(* IEC 61131-3 sources: plc-workbench/customers/naidis-metall/magazine-swivel/plc/src, 2 files *)

(* ---- plant_sim.st ---- *)
(* Plant model of the magazine and swivel station, for the sim target only.
   Reads the valve coils and writes the sensors, once per 10 ms scan before Station.
   Positions count scans: one count per scan, so 40 counts = 400 ms of travel. *)

PROGRAM PlantSim
    VAR_EXTERNAL
        MAG_CylExtended : BOOL;
        MAG_CylRetracted : BOOL;
        GRP_PartGripped : BOOL;
        SWV_AtPickup : BOOL;
        SWV_AtDropdown : BOOL;
        MAG_PickupOccupied : BOOL;
        MAG_CylRetract : BOOL;
        GRP_Grip : BOOL;
        GRP_Release : BOOL;
        SWV_ToPickup : BOOL;
        SWV_ToDropdown : BOOL;
        SIM_PartsInMagazine : INT;
        SIM_PartsDelivered : INT;
        SIM_PartsLost : INT;
        SIM_VacuumFault : BOOL;
        SIM_SwivelJam : BOOL;
        SIM_SorterBlocked : BOOL;
        LNK_NextReady : BOOL;
    END_VAR
    VAR CONSTANT
        MagStroke : INT := 40;    (* 0 = extended, MagStroke = retracted *)
        SwvStroke : INT := 50;    (* 0 = at dropdown, SwvStroke = at pickup *)
        SortScans : INT := 100;   (* the sorter takes a delivered part away in 1 s *)
    END_VAR
    VAR
        MagPos : INT := 0;
        SwvPos : INT := 0;
        PartInFront : BOOL;       (* dropped from the magazine in front of the retracted cylinder *)
        PartAtPickup : BOOL;
        PartOnGripper : BOOL;
        Vacuum : BOOL;
        VacuumBuildUp : TON;
        SortCount : INT := 0;     (* > 0 while the sorter is busy with the last part *)
    END_VAR

    (* 1A1 magazine cylinder: 5/2 single solenoid, coil on retracts, spring extends *)
    IF MAG_CylRetract THEN
        IF MagPos < MagStroke THEN MagPos := MagPos + 1; END_IF;
    ELSIF MagPos > 0 THEN
        MagPos := MagPos - 1;
    END_IF;
    IF MagPos = MagStroke AND NOT PartInFront AND SIM_PartsInMagazine > 0 THEN
        PartInFront := TRUE;
        SIM_PartsInMagazine := SIM_PartsInMagazine - 1;
    END_IF;
    IF MagPos = 0 AND PartInFront THEN
        PartInFront := FALSE;
        PartAtPickup := TRUE;
    END_IF;

    (* 3A1 swivel: 5/3 closed centre, stops with both coils off or both on *)
    IF NOT SIM_SwivelJam THEN
        IF SWV_ToPickup AND NOT SWV_ToDropdown AND SwvPos < SwvStroke THEN
            SwvPos := SwvPos + 1;
        ELSIF SWV_ToDropdown AND NOT SWV_ToPickup AND SwvPos > 0 THEN
            SwvPos := SwvPos - 1;
        END_IF;
    END_IF;

    (* 2A1 vacuum gripper: valve keeps its last coil *)
    IF GRP_Grip AND NOT GRP_Release THEN
        Vacuum := TRUE;
    ELSIF GRP_Release AND NOT GRP_Grip THEN
        Vacuum := FALSE;
    END_IF;
    IF Vacuum AND SwvPos = SwvStroke AND PartAtPickup THEN
        PartAtPickup := FALSE;
        PartOnGripper := TRUE;
    END_IF;
    IF PartOnGripper AND (NOT Vacuum OR SIM_VacuumFault) THEN
        PartOnGripper := FALSE;
        IF SwvPos = 0 AND LNK_NextReady THEN
            SIM_PartsDelivered := SIM_PartsDelivered + 1;
            SortCount := SortScans;
        ELSIF SwvPos = 0 THEN
            SIM_PartsLost := SIM_PartsLost + 1;      (* dropped onto a sorter that was not ready *)
        ELSIF SwvPos = SwvStroke THEN
            PartAtPickup := TRUE;
        ELSE
            SIM_PartsLost := SIM_PartsLost + 1;
        END_IF;
    END_IF;
    VacuumBuildUp(IN := Vacuum AND PartOnGripper, PT := T#100MS);

    (* colour sorter downstream: ready over the IR link unless busy or blocked *)
    IF SortCount > 0 THEN SortCount := SortCount - 1; END_IF;

    MAG_CylExtended := MagPos = 0;
    MAG_CylRetracted := MagPos = MagStroke;
    MAG_PickupOccupied := PartAtPickup;
    SWV_AtDropdown := SwvPos = 0;
    SWV_AtPickup := SwvPos = SwvStroke;
    GRP_PartGripped := VacuumBuildUp.Q;
    LNK_NextReady := SortCount = 0 AND NOT SIM_SorterBlocked;
END_PROGRAM

(* ---- station.st ---- *)
(* Magazine and swivel station: step sequence.
   Spec: ../magazine-swivel.spec.md, section 5.
   I/O symbols are globals declared by the target (targets/*.st). *)

TYPE
    StepT : (
        S0_Ready,
        S1_MagRetract,
        S2_MagPushOut,
        S3_SwvToPickup,
        S4_VacuumOn,
        S5_WaitNextReady,
        S6_SwvToDropdown,
        S7_VacuumOff,
        S8_CycleEnd,
        S9_MagEmpty,
        S90_HomingRequired,
        S91_HomeSwivel,
        S92_HomeVacuumOff,
        S99_Alarm);
END_TYPE

PROGRAM Station
    VAR_EXTERNAL
        PNL_StartButton : BOOL;
        PNL_StopReleased : BOOL;
        PNL_Manual : BOOL;
        PNL_ResetButton : BOOL;
        PNL_EStopOk : BOOL;
        MAG_CylExtended : BOOL;
        MAG_CylRetracted : BOOL;
        GRP_PartGripped : BOOL;
        SWV_AtPickup : BOOL;
        SWV_AtDropdown : BOOL;
        MAG_PickupOccupied : BOOL;
        LNK_NextReady : BOOL;
        PNL_StartLamp : BOOL;
        PNL_ResetLamp : BOOL;
        PNL_LampQ1 : BOOL;
        PNL_LampQ2 : BOOL;
        MAG_CylRetract : BOOL;
        GRP_Grip : BOOL;
        GRP_Release : BOOL;
        SWV_ToPickup : BOOL;
        SWV_ToDropdown : BOOL;
        StepNo : INT;   (* Step as a number (S90 = 90) for HMI and simulation *)
    END_VAR
    VAR
        CurStep : StepT := S90_HomingRequired;
        LastStep : StepT := S90_HomingRequired;
        StepTimer : TON;
        StepTime : TIME;
        FirstScan : BOOL := TRUE;
        StartTrig : R_TRIG;
        ResetTrig : R_TRIG;
        StartP : BOOL;
        ResetP : BOOL;
        BlinkTimer : TON;
        Blink1Hz : BOOL;
        Home : BOOL;
        StopReq : BOOL;
    END_VAR

    StepTimer(IN := CurStep = LastStep, PT := T#24H);  (* restarts on every step change *)
    StepTime := StepTimer.ET;
    LastStep := CurStep;

    BlinkTimer(IN := NOT BlinkTimer.Q, PT := T#500MS);
    IF BlinkTimer.Q THEN Blink1Hz := NOT Blink1Hz; END_IF;

    StartTrig(CLK := PNL_StartButton);
    StartP := StartTrig.Q;
    ResetTrig(CLK := PNL_ResetButton);
    ResetP := ResetTrig.Q;

    Home := MAG_CylExtended AND SWV_AtDropdown;

    IF CurStep = S0_Ready OR CurStep = S9_MagEmpty THEN
        StopReq := FALSE;
    ELSIF NOT PNL_StopReleased THEN
        StopReq := TRUE;
    END_IF;

    IF FirstScan THEN
        IF Home THEN CurStep := S0_Ready; ELSE CurStep := S90_HomingRequired; END_IF;
    ELSIF NOT PNL_EStopOk THEN
        CurStep := S90_HomingRequired;
    ELSE
        CASE CurStep OF
        S90_HomingRequired:
            IF ResetP AND PNL_EStopOk THEN CurStep := S91_HomeSwivel; END_IF;

        S91_HomeSwivel:
            IF SWV_AtDropdown THEN CurStep := S92_HomeVacuumOff;
            ELSIF StepTime >= T#3S THEN CurStep := S99_Alarm; END_IF;

        S92_HomeVacuumOff:
            IF StepTime >= T#50MS AND Home THEN CurStep := S0_Ready;
            ELSIF StepTime >= T#3S THEN CurStep := S99_Alarm; END_IF;

        S0_Ready:
            IF NOT Home THEN CurStep := S90_HomingRequired;
            ELSIF StartP AND PNL_StopReleased THEN
                IF MAG_PickupOccupied THEN CurStep := S3_SwvToPickup; ELSE CurStep := S1_MagRetract; END_IF;
            END_IF;

        S1_MagRetract:
            IF MAG_CylRetracted THEN CurStep := S2_MagPushOut;
            ELSIF StepTime >= T#3S THEN CurStep := S99_Alarm; END_IF;

        S2_MagPushOut:
            IF MAG_CylExtended THEN
                IF MAG_PickupOccupied THEN CurStep := S3_SwvToPickup; ELSE CurStep := S9_MagEmpty; END_IF;
            ELSIF StepTime >= T#3S THEN CurStep := S99_Alarm; END_IF;

        S3_SwvToPickup:
            IF SWV_AtPickup THEN CurStep := S4_VacuumOn;
            ELSIF StepTime >= T#3S THEN CurStep := S99_Alarm; END_IF;

        S4_VacuumOn:
            IF GRP_PartGripped THEN CurStep := S5_WaitNextReady;
            ELSIF StepTime >= T#3S THEN CurStep := S99_Alarm; END_IF;  (* part not gripped *)

        S5_WaitNextReady:
            IF NOT GRP_PartGripped THEN CurStep := S99_Alarm;          (* part lost *)
            ELSIF LNK_NextReady THEN CurStep := S6_SwvToDropdown; END_IF;

        S6_SwvToDropdown:
            IF NOT GRP_PartGripped THEN CurStep := S99_Alarm;          (* part lost *)
            ELSIF SWV_AtDropdown THEN CurStep := S7_VacuumOff;
            ELSIF StepTime >= T#3S THEN CurStep := S99_Alarm; END_IF;

        S7_VacuumOff:
            IF StepTime >= T#50MS THEN CurStep := S8_CycleEnd; END_IF;

        S8_CycleEnd:
            IF StopReq OR PNL_Manual THEN CurStep := S0_Ready; ELSE CurStep := S1_MagRetract; END_IF;

        S9_MagEmpty:
            IF NOT Home THEN CurStep := S90_HomingRequired;
            ELSIF StartP AND PNL_StopReleased THEN CurStep := S1_MagRetract; END_IF;

        S99_Alarm:
            IF ResetP AND PNL_EStopOk THEN CurStep := S91_HomeSwivel; END_IF;
        END_CASE;
    END_IF;

    (* one line per output; never assigned anywhere else *)
    MAG_CylRetract := CurStep = S1_MagRetract AND SWV_AtDropdown;
    GRP_Grip := CurStep = S4_VacuumOn OR CurStep = S5_WaitNextReady OR CurStep = S6_SwvToDropdown;
    GRP_Release := CurStep = S92_HomeVacuumOff OR CurStep = S7_VacuumOff;
    SWV_ToPickup := (CurStep = S3_SwvToPickup OR CurStep = S4_VacuumOn OR CurStep = S5_WaitNextReady)
        AND MAG_CylExtended;
    SWV_ToDropdown := CurStep = S91_HomeSwivel OR CurStep = S92_HomeVacuumOff
        OR CurStep = S6_SwvToDropdown OR CurStep = S7_VacuumOff;
    PNL_StartLamp := (CurStep = S0_Ready OR CurStep = S9_MagEmpty) AND Blink1Hz
        OR CurStep = S1_MagRetract OR CurStep = S2_MagPushOut OR CurStep = S3_SwvToPickup
        OR CurStep = S4_VacuumOn OR CurStep = S5_WaitNextReady OR CurStep = S6_SwvToDropdown
        OR CurStep = S7_VacuumOff OR CurStep = S8_CycleEnd;
    PNL_ResetLamp := CurStep = S90_HomingRequired AND (Blink1Hz OR NOT PNL_EStopOk)
        OR CurStep = S91_HomeSwivel OR CurStep = S92_HomeVacuumOff
        OR CurStep = S99_Alarm AND Blink1Hz;
    PNL_LampQ1 := PNL_ResetLamp;   (* same steps and modifiers as the reset lamp *)
    PNL_LampQ2 := PNL_ResetLamp OR CurStep = S9_MagEmpty AND Blink1Hz;

    CASE CurStep OF
    S0_Ready: StepNo := 0;
    S1_MagRetract: StepNo := 1;
    S2_MagPushOut: StepNo := 2;
    S3_SwvToPickup: StepNo := 3;
    S4_VacuumOn: StepNo := 4;
    S5_WaitNextReady: StepNo := 5;
    S6_SwvToDropdown: StepNo := 6;
    S7_VacuumOff: StepNo := 7;
    S8_CycleEnd: StepNo := 8;
    S9_MagEmpty: StepNo := 9;
    S90_HomingRequired: StepNo := 90;
    S91_HomeSwivel: StepNo := 91;
    S92_HomeVacuumOff: StepNo := 92;
    S99_Alarm: StepNo := 99;
    END_CASE;

    FirstScan := FALSE;
END_PROGRAM
